(* IEC 61131-3 sources: tsplc/examples/bottling-line/raw-st/src, 1 file *)

(* ---- Main.st ---- *)
PROGRAM Main
VAR
	Capper : FB_Capper;
END_VAR
PRG_ReadInputs();
PRG_Transport();
Capper(BottlePresent := IO.BottlePresent);
IO.CapperRun := Capper.Running;
PRG_Publish();
END_PROGRAM
